// TIA Portal V20 export
// export: Created 2026-10-19T18:45:09.0304786Z, ExportSetting None, DisplayName Totally Integrated Automation Portal, DisplayVersion V20 Update 6, DisplayName TIA Portal Openness, DisplayVersion V20 Update 6, DisplayName TIA Portal Version Control Interface, DisplayVersion V20 Update 6, DisplayName SINAMICS Startdrive Advanced, DisplayVersion V20 SP1, DisplayName SINAMICS Startdrive G130, G150, S120, S150, SINAMICS MV, G220, S200, S210, DisplayVersion V20 SP1, DisplayName SINAMICS Startdrive G110M, G120, G120C, G120D, G120P, G115D, DisplayVersion V20 SP1, DisplayName STEP 7 Professional, DisplayVersion V20 Update 6, DisplayName STEP 7 Safety, DisplayVersion V20 Update 2, DisplayName WinCC Basic/Comfort/Advanced, DisplayVersion V20 Update 6, DisplayName WinCC Unified, DisplayVersion V20 Update 6
VAR_GLOBAL   // PLC tag table "CNV_HMI"
   "Manual_Sfty_Stopper_Up(1)" AT %M8.5 : Bool;
   "Manual_Sfty_Stopper_Down(1)" AT %M8.7 : Bool;
   CNV_ID_HMI AT %MD1125 : DInt;
   Manual_Bwd_HMI AT %M4.2 : Bool;
   "Reset_HMI(1)" AT %M4.5 : Bool;
   Manual_Fwd_HMI AT %M4.1 : Bool;
   Enable_HMI AT %M2.7 : Bool;
   CNV_ID_HMI_Old AT %MD72 : DInt;
   "Enable_HMI(1)" AT %M20.1 : Bool;
   "Transfer_To_ID_HMI(1)" AT %MD29 : DInt;
   "Manual_Bwd_HMI(1)" AT %M6.1 : Bool;
   Reset_HMI AT %M3.0 : Bool;
   Stop_HMI AT %M2.6 : Bool;
   "Start_Transfer_HMI(1)" AT %M5.3 : Bool;
   Start_Transfer_HMI AT %M3.6 : Bool;
   "CNV_ID_HMI(1)" AT %MD1133 : DInt;
   "Transfer_From_ID_HMI(1)" AT %MD1151 : DInt;
   "Manual_Fwd_HMI(1)" AT %M6.0 : Bool;
   Mode_Change_HMI AT %MW1129 : UInt;
   Transfer_To_ID_HMI AT %MD15 : DInt;
   "Mode_Change_HMI(1)" AT %MW21 : UInt;
   Transfer_From_ID_HMI AT %MD1147 : DInt;
   "CNV_ID_HM_Old(1)" AT %MD76 : DInt;
   "CNV_In_Out(1)" AT %M80.1 : Bool;
   CNV_Level_Selected_OLD AT %MW122 : UInt;
   "Cnv_Occupied_HMI(1)" AT %M7.7 : Bool;
   Mode_HMI AT %MW33 : UInt;
   "Running_HMI(1)" AT %M7.5 : Bool;
   "Enabled_HMI(1)" AT %M7.2 : Bool;
   Motor_Speed_Actual_HMI AT %MW50 : UInt;
   Running_HMI AT %M6.6 : Bool;
   "SM_State_HMI(1)" AT %MW62 : UInt;
   "Warning_HMI(1)" AT %MW54 : UInt;
   Stopped_HMI AT %M6.5 : Bool;
   Enabled_HMI AT %M6.3 : Bool;
   Error_HMI AT %M6.4 : Bool;
   "Motor_Speed_Requested_HMI(1)" AT %MW66 : UInt;
   "Mode_HMI(1)" AT %MW52 : UInt;
   Warning_HMI AT %MW35 : UInt;
   "Stopped_HMI(1)" AT %M7.4 : Bool;
   Motor_Direction_HMI AT %MW46 : UInt;
   SM_State_HMI AT %MW44 : UInt;
   "Ready_For_Task_HMI(1)" AT %M7.6 : Bool;
   Ready_For_Task_HMI AT %M6.7 : Bool;
   Cnv_Occupied_HMI AT %M7.0 : Bool;
   "Error_HMI(1)" AT %M7.3 : Bool;
   Motor_Speed_Requested_HMI AT %MW48 : UInt;
   "Motor_Direction_HMI(1)" AT %MW64 : UInt;
   "Motor_Speed_Actual_HMI(1)" AT %MW68 : UInt;
   CNV_Motor_Ready AT %M60.0 : Bool;
   "CNV_Motor_Current_Actual_HMI(1)" AT %MD142 : Real;
   CNV_Motor_Status_HMI AT %MW124 : UInt;
   "CNV_Motor_Status_HMI(1)" AT %MW126 : UInt;
   CNV_Motor_Current_Actual_HMI AT %MD138 : Real;
   "CNV_Motor_Ready(1)" AT %M60.1 : Bool;
   CNV_Level_Selected AT %MW146 : UInt;
   CNV_System_Selected AT %MW150 : UInt;
   "UpDown(1)" AT %MW84 : UInt;
   CNV_Motor_Actual_Torque AT %MD170 : Real;
   "CNV_Motor_Actual_Torque(1)" AT %MD178 : Real;
   HMI_Light_Guard_Bypass AT %M186.1 : Bool;
   "Light_Guard_Bypass(1)" AT %M186.4 : Bool;
   "Light_Guard_Bypass(2)" AT %M186.2 : Bool;
   CVTD_CNV2_Selected AT %MW106 : UInt;
END_VAR
